# EPICS substitutions: iocs/motor/npoint-ioc/db/C300.substitutions
# C's iocNPoint C300.substitutions, P and PORT from st.cmd.
file "$(MOTOR)/db/asyn_motor.db"
{
pattern
{N,  M,       DTYP,         ADDR,  DESC,          EGU,  DIR,  VELO,  VBAS,  ACCL,  BDST,  BVEL,  BACC,  MRES,             PREC,  DHLM,  DLLM,   INIT}
{1,  "m$(N)", "asynMotor",  0,     "motor $(N)",  um,   Pos,  1,     .1,    .2,    0,     1,     .2,    9.5367431641e-5,  5,     50,    -50,    ""}
{2,  "m$(N)", "asynMotor",  1,     "motor $(N)",  um,   Pos,  1,     .1,    .2,    0,     1,     .2,    9.5367431641e-5,  5,     50,    -50,    ""}
{3,  "m$(N)", "asynMotor",  2,     "motor $(N)",  um,   Pos,  1,     .1,    .2,    0,     1,     .2,    2.384185791e-5,   5,     12.5,  -12.5,  ""}
}
